(* IEC 61131-3 sources: PortalRobot/Portal_robot/Device/application/FB (part 6) *)

(* ---- FB_TWO_PALLET.st ---- *)
FUNCTION_BLOCK FB_TWO_PALLET
VAR_INPUT
	xSelected : BOOL;
	xManual : BOOL;
	xSafe : BOOL;
	xRobotSwapWindow : BOOL; // Завершено последнее обслуживание: разрешён автоматический обмен
	xRobotOperation : BOOL; // Текущая или уже выданная операция с этим магазином
	xPointsConfigured : BOOL; // Собственная база магазина нужна для ввода в автомат
	xRobotGeometryReady : BOOL; // Собственная база магазина и поддерживаемый интерфейс робота
	xRobotMagazineReady : BOOL; // Ошибки и геометрия магазина; содержимое не блокирует включение
	xConnection : BOOL; // Heartbeat HMI нужен только для ручных команд
	xStopRequest : BOOL; // Общий Stop прерывает движение, но не отключает неподвижный магазин
	xAutoSwap : BOOL;
	xOtherLoaded : BOOL;
	xActivePalletEditAllowed : BOOL;
	xConfigurationChanged : BOOL;
    xIoPneumaticOverride : BOOL; // Прямое воздействие на катушки снимает подтверждение расстановки
	xExternalCommandRejected : BOOL;
	Command : ST_TWO_PALLET_COMMAND;
	Config : ST_TWO_PALLET_CONFIG;
	Input : ST_TWO_PALLET_INPUT;
END_VAR
VAR_OUTPUT
	Status : ST_TWO_PALLET_STATUS;
	Diag : ST_TWO_PALLET_DIAG;
	Error : ST_TWO_PALLET_ERRORS;
	Output : ST_TWO_PALLET_OUTPUT;
END_VAR
VAR
	ePreviousState : E_TWO_PALLET_STATE := E_TWO_PALLET_STATE.IDLE;
	uiFrom : UINT;
	uiTo : UINT;
	uiSelected : UINT;
	uiCandidate : UINT;
	uiPreviousCandidate : UINT;
	uiConfirmedCandidate : UINT;
	uiManualSelected : UINT;
	uiJogDirection : UINT;
	uiSignals : UINT;
	uiSelectedSignals : UINT;
	uiTargetSignals : UINT;
	xPreviousBaseValid : BOOL;
	xConfigValid : BOOL;
	xContradiction : BOOL;
	xPairValid : BOOL;
	xWork : BOOL;
	xExchange : BOOL;
	xIdle : BOOL;
	xBase : BOOL;
	xManualSetupAllowed : BOOL;
	xRecovery : BOOL;
	xPneumaticBase : BOOL;
	xPneumaticRecovery : BOOL;
	xManualPneumaticState : BOOL;
	xAutomaticState : BOOL;
	xAxisMotionState : BOOL;
	xManualState : BOOL;
	xEnableBaseAllowed : BOOL;
	xAutoSwapAllowed : BOOL;
	xExchangeStartedManual : BOOL; // Обмен начат в ручном режиме: без проверки роботной зоны/точек
	xCommandPresent : BOOL;
	xAccepted : BOOL;
	xStateEntry : BOOL;
	xSeenMotion : BOOL;
	xSeenDone : BOOL;
	xLiftUpCommand : BOOL;
	xLiftDownCommand : BOOL;
	xSelectCommand : BOOL;
	xManualLockCommand : BOOL;
	xManualStopCommand : BOOL;
	xManualLockOutTarget : BOOL;
	xManualStopOutTarget : BOOL;
	xLockOutTarget : BOOL;
	xStopOutTarget : BOOL;
	xStartupInitialized : BOOL;
	xTrustedAtScanStart : BOOL;
	lrWork : LREAL;
	lrTarget : LREAL;
	lrSpan : LREAL;
	rTravel : REAL;
	tStateLimit : TIME;
	tonState : TON;
	tonCoil : TON;
	tonJogLease : TON;
	dwPreviousError : DWORD;
END_VAR
VAR CONSTANT
	ERR_DRIVE : DWORD := DWORD#16#100;
	ERR_SENSOR_CONTRADICTION : DWORD := DWORD#16#200;
	ERR_CYLINDER_TIMEOUT : DWORD := DWORD#16#400;
	ERR_MOTION_TIMEOUT : DWORD := DWORD#16#800;
	ERR_LOGIC : DWORD := DWORD#16#1000;
	ERR_SEQUENCE_INTERRUPTED : DWORD := DWORD#16#2000;
	WRN_COMMAND_REJECTED : UINT := UINT#30;
	WRN_ENABLE_POINTS : UINT := UINT#18; // Общий код с FB_MAGAZINE для отсутствующей базы
	WRN_START_REJECTED_BY_OPERATOR : UINT := UINT#31;
	JOG_POSITIVE : UINT := UINT#1;
	JOG_NEGATIVE : UINT := UINT#2;
END_VAR

// --- BEGIN IMPLEMENTATION ---

// Шаги, разрешения и подтверждение положения не восстанавливаются после старта PLC.
IF NOT xStartupInitialized THEN
	Diag.eState := E_TWO_PALLET_STATE.IDLE;
	ePreviousState := E_TWO_PALLET_STATE.IDLE;
	Status.xConfirmed := FALSE;
	Status.xEnabled := FALSE;
	xStartupInitialized := TRUE;
END_IF;

Status.xCompleted := FALSE;
Status.Input := Input;
xTrustedAtScanStart := Status.xConfirmed;

// Все выходные команды импульсные или формируются заново на каждом скане.
Output.xPowerOn := FALSE;
Output.xPowerOff := FALSE;
Output.xDriveReset := FALSE;
Output.xHome := FALSE;
Output.xMove := FALSE;
Output.xStop := FALSE;
Output.xJogPositive := FALSE;
Output.xJogNegative := FALSE;
Output.xTeachOperator := FALSE;
Output.xTeachWork := FALSE;
xLiftUpCommand := FALSE;
xLiftDownCommand := FALSE;
xSelectCommand := FALSE;
xManualLockCommand := FALSE;
xManualStopCommand := FALSE;

// Конфигурация механизма.
xConfigValid := Config.xConfigured
	AND Config.xSignalPatternsConfigured
	AND IsSignalConfigurationValid(uiP1Signals := Config.uiP1Signals, uiP2Signals := Config.uiP2Signals)
	AND (Config.lrTolerance > 0.0)
	AND (Config.lrTolerance <= 20.0)
	AND (ABS(Config.lrWorkP1 - Config.lrExchange) > 2.0 * Config.lrTolerance)
	AND (ABS(Config.lrWorkP2 - Config.lrExchange) > 2.0 * Config.lrTolerance)
	AND ((Config.lrWorkP1 - Config.lrExchange) * (Config.lrWorkP2 - Config.lrExchange) > 0.0)
	AND (Config.lrVelocity > 0.0)
	AND (Config.lrAcceleration > 0.0)
	AND (Config.lrDeceleration > 0.0)
	AND (Config.lrJerk > 0.0)
	AND (Config.tPulse >= T#50MS)
	AND (Config.tCylinder > Config.tPulse)
	AND (Config.tMove > T#0S)
	AND (Config.tHome > T#0S);
Status.xConfigValid := xConfigValid;

// Фактическое состояние пневматики и каретки.
xContradiction := (Input.xLiftUp AND Input.xLiftDown)
	OR (Input.xLockIn AND Input.xLockOut)
	OR (Input.xStopIn AND Input.xStopOut)
	OR (Input.xLimitNegative AND Input.xLimitPositive);
xPairValid := (Input.xLockIn XOR Input.xLockOut)
	AND (Input.xStopIn XOR Input.xStopOut);

uiSignals := UINT#0;
IF Input.xLiftDown THEN uiSignals := uiSignals OR UINT#1; END_IF;
IF Input.xLiftUp THEN uiSignals := uiSignals OR UINT#2; END_IF;
IF Input.xLockIn THEN uiSignals := uiSignals OR UINT#4; END_IF;
IF Input.xLockOut THEN uiSignals := uiSignals OR UINT#8; END_IF;
IF Input.xStopIn THEN uiSignals := uiSignals OR UINT#16; END_IF;
IF Input.xStopOut THEN uiSignals := uiSignals OR UINT#32; END_IF;

uiSelected := UINT#0;
IF xPairValid THEN
	IF (uiSignals AND UINT#60) = (Config.uiP1Signals AND UINT#60) THEN
		uiSelected := UINT#1;
	ELSIF (uiSignals AND UINT#60) = (Config.uiP2Signals AND UINT#60) THEN
		uiSelected := UINT#2;
	END_IF;
END_IF;
xPairValid := xPairValid AND (uiSelected <> UINT#0);

lrWork := Config.lrWorkP1;
uiSelectedSignals := Config.uiP1Signals;
IF uiSelected = UINT#2 THEN
	lrWork := Config.lrWorkP2;
	uiSelectedSignals := Config.uiP2Signals;
END_IF;

xWork := xConfigValid
	AND Input.xHomed
	AND Input.xStandstill
	AND xPairValid
	AND (ABS(Input.lrPosition - lrWork) <= Config.lrTolerance);
xExchange := xConfigValid
	AND Input.xHomed
	AND Input.xStandstill
	AND (ABS(Input.lrPosition - Config.lrExchange) <= Config.lrTolerance);

uiCandidate := UINT#0;
IF xWork
	AND (uiSignals = uiSelectedSignals)
	AND NOT xContradiction
	AND NOT Input.xDriveError
	AND NOT Status.xHomeRequired THEN
	uiCandidate := uiSelected;
END_IF;

xIdle := Diag.eState = E_TWO_PALLET_STATE.IDLE;
xAutomaticState := (Diag.eState = E_TWO_PALLET_STATE.AUTO_LOWER)
	OR (Diag.eState = E_TWO_PALLET_STATE.AUTO_MOVE_TO_EXCHANGE)
	OR (Diag.eState = E_TWO_PALLET_STATE.AUTO_SELECT_PALLET)
	OR (Diag.eState = E_TWO_PALLET_STATE.AUTO_MOVE_TO_WORK)
	OR (Diag.eState = E_TWO_PALLET_STATE.AUTO_RAISE);
xAxisMotionState := (Diag.eState = E_TWO_PALLET_STATE.AUTO_MOVE_TO_EXCHANGE)
	OR (Diag.eState = E_TWO_PALLET_STATE.AUTO_MOVE_TO_WORK)
	OR (Diag.eState = E_TWO_PALLET_STATE.MANUAL_MOVE)
	OR (Diag.eState = E_TWO_PALLET_STATE.MANUAL_HOME)
	OR (Diag.eState = E_TWO_PALLET_STATE.MANUAL_JOG);
xManualState := (Diag.eState = E_TWO_PALLET_STATE.MANUAL_LOWER)
	OR (Diag.eState = E_TWO_PALLET_STATE.MANUAL_RAISE)
	OR (Diag.eState = E_TWO_PALLET_STATE.MANUAL_SELECT_PALLET)
	OR (Diag.eState = E_TWO_PALLET_STATE.MANUAL_MOVE)
	OR (Diag.eState = E_TWO_PALLET_STATE.MANUAL_HOME)
	OR (Diag.eState = E_TWO_PALLET_STATE.MANUAL_JOG)
	OR (Diag.eState = E_TWO_PALLET_STATE.MANUAL_LOCK)
	OR (Diag.eState = E_TWO_PALLET_STATE.MANUAL_STOP);
xManualPneumaticState := (Diag.eState = E_TWO_PALLET_STATE.MANUAL_LOWER)
	OR (Diag.eState = E_TWO_PALLET_STATE.MANUAL_LOCK)
	OR (Diag.eState = E_TWO_PALLET_STATE.MANUAL_STOP);

xBase := xSelected
	AND xConfigValid
	AND Input.xIoMapped
	AND Input.xAxisBound
	AND xSafe
	AND NOT xRobotOperation;
xManualSetupAllowed := xManual
	AND NOT Status.xEnabled
	AND NOT xRobotOperation;
xRecovery := xBase
	AND xManualSetupAllowed
	AND xConnection
	AND xIdle
	AND Input.xStandstill;
xPneumaticBase := xSelected
	AND xManualSetupAllowed
	AND xSafe
	AND Input.xIoMapped
	AND Input.xStandstill;
xPneumaticRecovery := xPneumaticBase AND xIdle;

Status.uiCandidate := uiCandidate;
Status.uiSelected := uiSelected;

// Любое изменение достоверной расстановки аннулирует старое подтверждение.
IF (uiCandidate <> uiPreviousCandidate) OR (xBase <> xPreviousBaseValid) THEN
	Status.udiRevision := Status.udiRevision + UDINT#1;
	IF Status.udiRevision = UDINT#0 THEN
		Status.udiRevision := UDINT#1;
	END_IF;
END_IF;
uiPreviousCandidate := uiCandidate;
xPreviousBaseValid := xBase;

IF xConfigurationChanged THEN
	Status.xConfirmed := FALSE;
	Status.xEnabled := FALSE;
	Status.udiRevision := Status.udiRevision + UDINT#1;
	IF Status.udiRevision = UDINT#0 THEN
		Status.udiRevision := UDINT#1;
	END_IF;
END_IF;

IF xIoPneumaticOverride THEN
    Status.xConfirmed := FALSE;
    Status.xEnabled := FALSE;
    Status.udiRevision := Status.udiRevision + UDINT#1;
    IF Status.udiRevision = UDINT#0 THEN Status.udiRevision := UDINT#1; END_IF;
END_IF;

IF NOT xSelected
	OR NOT xSafe
	OR NOT Input.xAxisBound
	OR NOT Input.xIoMapped
	OR NOT xConfigValid
	OR Input.xDriveError
	OR NOT Input.xPowered
	OR (xIdle AND (uiCandidate <> uiConfirmedCandidate)) THEN
	Status.xConfirmed := FALSE;
END_IF;
// Первая невыполненная предпосылка для HMI.
Diag.uiReason := UINT#0;
IF NOT xSelected THEN
	Diag.uiReason := UINT#1;
ELSIF NOT xConfigValid THEN
	Diag.uiReason := UINT#2;
ELSIF NOT Input.xAxisBound OR NOT Input.xIoMapped THEN
	Diag.uiReason := UINT#3;
ELSIF NOT xSafe THEN
	Diag.uiReason := UINT#4;
ELSIF NOT xConnection THEN
	Diag.uiReason := UINT#17;
ELSIF Input.xDriveError THEN
	Diag.uiReason := UINT#6;
ELSIF Error.dwErrorActive <> DWORD#0 THEN
	Diag.uiReason := UINT#19;
ELSIF NOT Input.xPowered THEN
	Diag.uiReason := UINT#18;
ELSIF xContradiction THEN
	Diag.uiReason := UINT#7;
ELSIF Status.xHomeRequired OR NOT Input.xHomed THEN
	Diag.uiReason := UINT#8;
ELSIF NOT xPairValid THEN
	Diag.uiReason := UINT#9;
ELSIF NOT Input.xStandstill THEN
	Diag.uiReason := UINT#10;
ELSIF NOT xWork THEN
	Diag.uiReason := UINT#11;
ELSIF uiSignals <> uiSelectedSignals THEN
	Diag.uiReason := UINT#12;
ELSIF NOT xIdle THEN
	Diag.uiReason := UINT#22;
ELSIF xRobotOperation THEN
	Diag.uiReason := UINT#5;
ELSIF xManual AND Status.xEnabled THEN
	Diag.uiReason := UINT#21;
ELSIF NOT xManual AND NOT xRobotSwapWindow THEN
	Diag.uiReason := UINT#23;
ELSIF NOT xRobotMagazineReady THEN
	Diag.uiReason := UINT#16;
ELSIF NOT xPointsConfigured THEN
	Diag.uiReason := UINT#15;
ELSIF NOT Status.xConfirmed AND NOT xManual THEN
	Diag.uiReason := UINT#20;
ELSIF NOT Status.xConfirmed THEN
	Diag.uiReason := UINT#13;
END_IF;

// Аварии механизма: биты 8..13 зарезервированы в MAGAZINE_LOGIC_1/2.
IF xSelected AND Input.xDriveError THEN
	Error.dwErrorActive := Error.dwErrorActive OR ERR_DRIVE;
	Status.xHomeRequired := TRUE;
END_IF;

IF xSelected AND xContradiction THEN
	Error.dwErrorActive := Error.dwErrorActive OR ERR_SENSOR_CONTRADICTION;
END_IF;

IF xSelected
	AND NOT xIdle
	AND (((NOT xBase) AND NOT (xManualPneumaticState AND xPneumaticBase))
		OR (xManualState AND NOT xManual)
		OR ((NOT xConnection) AND xManualState AND NOT xManualPneumaticState) OR xStopRequest
		OR (xAutomaticState AND ((xExchangeStartedManual AND NOT xManual)
			OR (NOT xExchangeStartedManual AND NOT xRobotSwapWindow)))) THEN
	Error.dwErrorActive := Error.dwErrorActive OR ERR_SEQUENCE_INTERRUPTED;
	Diag.eState := E_TWO_PALLET_STATE.IDLE;
	Output.xStop := TRUE;
END_IF;

IF xSelected AND (xTrustedAtScanStart OR xAutomaticState) THEN
	IF ((Diag.eState <> E_TWO_PALLET_STATE.AUTO_SELECT_PALLET) AND NOT xPairValid)
		OR (((Diag.eState = E_TWO_PALLET_STATE.AUTO_MOVE_TO_EXCHANGE)
			OR (Diag.eState = E_TWO_PALLET_STATE.AUTO_MOVE_TO_WORK))
			AND (NOT Input.xLiftDown OR Input.xLiftUp))
		OR (xIdle AND (uiCandidate = UINT#0)) THEN
		Error.dwErrorActive := Error.dwErrorActive OR ERR_LOGIC;
	END_IF;
END_IF;

IF xSelected
	AND xTrustedAtScanStart
	AND (NOT xSafe
		OR NOT Input.xAxisBound
		OR NOT Input.xIoMapped
		OR NOT Input.xPowered) THEN
	Error.dwErrorActive := Error.dwErrorActive OR ERR_SEQUENCE_INTERRUPTED;
END_IF;

IF xSelected
	AND ((xContradiction AND NOT xIdle AND NOT xManualPneumaticState)
		OR (Input.xDriveError AND xAxisMotionState)) THEN
	Diag.eState := E_TWO_PALLET_STATE.IDLE;
	Output.xStop := TRUE;
END_IF;

IF xSelected AND NOT Input.xPowered AND (xAutomaticState OR xAxisMotionState) THEN
	Error.dwErrorActive := Error.dwErrorActive OR ERR_SEQUENCE_INTERRUPTED;
	Status.xHomeRequired := TRUE;
	Diag.eState := E_TWO_PALLET_STATE.IDLE;
	Output.xStop := TRUE;
END_IF;

IF Error.dwErrorActive <> DWORD#0 THEN
	Status.xEnabled := FALSE;
	Status.xConfirmed := FALSE;
	IF xAutomaticState THEN
		Diag.eState := E_TWO_PALLET_STATE.IDLE;
		Output.xStop := TRUE;
	END_IF;
END_IF;

// Разрешения считаются только владельцем механизма.
Status.xConfirmAllowed := xRecovery
	AND Input.xPowered
	AND (uiCandidate <> UINT#0)
	AND (Error.dwErrorActive = DWORD#0);
Status.xStartAllowed := Status.xConfirmAllowed
	AND xRobotMagazineReady
	AND xPointsConfigured;
// Включение подтверждённого магазина не двигает палету и не снимает резерв
// возврата изделия. Иначе Disable при грузе в роботе блокирует продолжение цикла.
// Общая технологическая готовность не зависит от heartbeat HMI.
xEnableBaseAllowed := xBase
	AND xIdle
	AND Status.xConfirmed
	AND xRobotMagazineReady
	AND xPointsConfigured
	AND (uiCandidate = Status.uiRobotPallet)
	AND Input.xPowered
	AND (Error.dwErrorActive = DWORD#0);
Status.xEnableAllowed := xEnableBaseAllowed AND xConnection;
// Обмен не требует глобальной остановки робота: проверяется только отсутствие
// текущей или уже выданной операции именно с этим магазином.
Status.xSwapAllowed := xBase
	AND xConnection
	AND xIdle
	AND Input.xStandstill
	AND Input.xPowered
	AND (Error.dwErrorActive = DWORD#0)
	AND Status.xConfirmed
	AND (uiCandidate = Status.uiRobotPallet)
	AND NOT Status.xEnabled
	AND NOT xStopRequest
	AND (xRobotSwapWindow OR xManual);
xAutoSwapAllowed := xEnableBaseAllowed
	AND xRobotSwapWindow
	AND Status.xEnabled
	AND xOtherLoaded;
Status.xPowerAllowed := xRecovery
	AND NOT Input.xDriveError
	AND NOT xContradiction;
Status.xDriveResetAllowed := xSelected
	AND xManualSetupAllowed
	AND xConnection
	AND Input.xAxisBound
	AND Input.xStandstill
	AND xIdle;
Status.xLowerAllowed := xPneumaticRecovery;
Status.xRaiseAllowed := xRecovery
	AND NOT xContradiction
	AND NOT Status.xHomeRequired;
Status.xSelectAllowed := xRecovery
	AND NOT xContradiction
	AND Input.xLiftDown
	AND NOT Input.xLiftUp
	AND xExchange;
// Наладочные команды замка и фиксатора независимы от подъёма и координаты.
// Это позволяет вернуть герконы в согласованное состояние после остановки.
Status.xLockAllowed := xPneumaticRecovery;
Status.xStopAllowed := xPneumaticRecovery;
Status.xHomeAllowed := xRecovery
	AND Input.xPowered
	AND NOT Input.xDriveError
	AND Input.xLiftDown
	AND NOT Input.xLiftUp
	AND xPairValid
	AND NOT xContradiction;
Status.xMoveAllowed := Status.xHomeAllowed
	AND Input.xHomed
	AND NOT Status.xHomeRequired;
Status.xJogAllowed := Status.xHomeAllowed;
Status.xTeachOperatorAllowed := Status.xMoveAllowed
	AND Input.xLiftDown
	AND NOT Input.xLiftUp;
Status.xTeachWorkAllowed := Status.xTeachOperatorAllowed
	AND ((uiSelected = UINT#1) OR (uiSelected = UINT#2));
Status.xResetAllowed := xRecovery
	AND (Error.dwErrorActive <> DWORD#0)
	AND NOT xContradiction
	AND NOT Input.xDriveError
	AND NOT Status.xHomeRequired
	AND xPairValid
	AND (Input.xLiftDown XOR Input.xLiftUp);
Status.xConfigAllowed := xSelected
	AND xManualSetupAllowed
	AND xIdle
	AND NOT Status.xEnabled
	AND (Input.xStandstill OR NOT Input.xAxisBound)
	AND NOT Input.xPowered;

// Командный интерфейс FB не зависит от транспортных номеров HMI 1..19.
xCommandPresent := Command.xEnable
	OR Command.xConfirm
	OR Command.xStart
	OR Command.xRejectStart
	OR Command.xDisable
	OR Command.xSwap
	OR Command.xPowerOn
	OR Command.xPowerOff
	OR Command.xDriveReset
	OR Command.xHome
	OR Command.xLower
	OR Command.xRaise
	OR Command.xSelectPallet
	OR Command.xLockIn
	OR Command.xLockOut
	OR Command.xStopIn
	OR Command.xStopOut
	OR Command.xMoveToExchange
	OR Command.xMoveToWork
	OR Command.xStop
	OR Command.xReset
	OR Command.xJogPositive
	OR Command.xJogNegative
	OR Command.xJogRelease
	OR Command.xTeachOperator
	OR Command.xTeachWork;
xAccepted := NOT xCommandPresent;

IF Command.xStart THEN
	IF Status.xStartAllowed
		AND (Command.udiRevision = Status.udiRevision)
		AND (Command.uiPallet = uiCandidate) THEN
		Status.uiRobotPallet := uiCandidate;
		uiConfirmedCandidate := uiCandidate;
		Status.xConfirmed := TRUE;
		Status.xEnabled := TRUE;
		Status.rP1 := 0.0;
		Status.rP2 := 0.0;
		IF uiCandidate = UINT#1 THEN
			Status.rP1 := 1.0;
		ELSE
			Status.rP2 := 1.0;
		END_IF;
		xAccepted := TRUE;
	END_IF;
ELSIF Command.xRejectStart THEN
	Diag.stWarning.uiCode := WRN_START_REJECTED_BY_OPERATOR;
	Diag.stWarning.udiSequence := Diag.stWarning.udiSequence + UDINT#1;
	IF Diag.stWarning.udiSequence = UDINT#0 THEN
		Diag.stWarning.udiSequence := UDINT#1;
	END_IF;
	xAccepted := TRUE;
ELSIF Command.xEnable THEN
	IF Status.xEnableAllowed THEN
		Status.xEnabled := TRUE;
		xAccepted := TRUE;
	END_IF;
ELSIF Command.xConfirm THEN
	IF Status.xConfirmAllowed
		AND (Command.udiRevision = Status.udiRevision)
		AND (Command.uiPallet = uiCandidate) THEN
		Status.uiRobotPallet := uiCandidate;
		uiConfirmedCandidate := uiCandidate;
		Status.xConfirmed := TRUE;
		Status.rP1 := 0.0;
		Status.rP2 := 0.0;
		IF uiCandidate = UINT#1 THEN
			Status.rP1 := 1.0;
		ELSE
			Status.rP2 := 1.0;
		END_IF;
		xAccepted := TRUE;
	END_IF;
ELSIF Command.xDisable THEN
	Status.xEnabled := FALSE;
	xAccepted := TRUE;
ELSIF Command.xSwap THEN
	IF Status.xSwapAllowed THEN
		xExchangeStartedManual := xManual;
		Diag.eState := E_TWO_PALLET_STATE.AUTO_LOWER;
		xAccepted := TRUE;
	END_IF;
ELSIF Command.xPowerOn THEN
	IF Status.xPowerAllowed THEN
		Output.xPowerOn := TRUE;
		xAccepted := TRUE;
	END_IF;
ELSIF Command.xPowerOff THEN
	IF Status.xDriveResetAllowed THEN
		Output.xPowerOff := TRUE;
		Status.xConfirmed := FALSE;
		Status.xEnabled := FALSE;
		xAccepted := TRUE;
	END_IF;
ELSIF Command.xDriveReset THEN
	IF Status.xDriveResetAllowed AND Input.xDriveError THEN
		Output.xDriveReset := TRUE;
		Status.xConfirmed := FALSE;
		Status.xEnabled := FALSE;
		Status.xHomeRequired := TRUE;
		xAccepted := TRUE;
	END_IF;
ELSIF Command.xHome THEN
	IF Status.xHomeAllowed THEN
		Diag.eState := E_TWO_PALLET_STATE.MANUAL_HOME;
		xAccepted := TRUE;
	END_IF;
ELSIF Command.xLower THEN
	IF Status.xLowerAllowed THEN
		Diag.eState := E_TWO_PALLET_STATE.MANUAL_LOWER;
		xAccepted := TRUE;
	END_IF;
ELSIF Command.xRaise THEN
	IF Status.xRaiseAllowed THEN
		Diag.eState := E_TWO_PALLET_STATE.MANUAL_RAISE;
		xAccepted := TRUE;
	END_IF;
ELSIF Command.xSelectPallet THEN
	IF Status.xSelectAllowed
		AND ((Command.uiPallet = UINT#1) OR (Command.uiPallet = UINT#2)) THEN
		uiTo := Command.uiPallet;
		Diag.eState := E_TWO_PALLET_STATE.MANUAL_SELECT_PALLET;
		xAccepted := TRUE;
	END_IF;
ELSIF Command.xLockIn OR Command.xLockOut THEN
	IF Status.xLockAllowed THEN
		xManualLockOutTarget := Command.xLockOut;
		Diag.eState := E_TWO_PALLET_STATE.MANUAL_LOCK;
		xAccepted := TRUE;
	END_IF;
ELSIF Command.xStopIn OR Command.xStopOut THEN
	IF Status.xStopAllowed THEN
		xManualStopOutTarget := Command.xStopOut;
		Diag.eState := E_TWO_PALLET_STATE.MANUAL_STOP;
		xAccepted := TRUE;
	END_IF;
ELSIF Command.xMoveToExchange OR Command.xMoveToWork THEN
	IF Status.xMoveAllowed THEN
		lrTarget := Config.lrExchange;
		IF Command.xMoveToWork THEN
			lrTarget := lrWork;
		END_IF;
		Diag.eState := E_TWO_PALLET_STATE.MANUAL_MOVE;
		xAccepted := TRUE;
	END_IF;
ELSIF Command.xStop THEN
	Status.xEnabled := FALSE;
	// Stop неподвижного механизма не является ручным вмешательством.
	IF (Diag.eState <> E_TWO_PALLET_STATE.IDLE) OR (Input.xPowered AND NOT Input.xStandstill) THEN
		Output.xStop := TRUE;
		Status.xConfirmed := FALSE;
		Error.dwErrorActive := Error.dwErrorActive OR ERR_SEQUENCE_INTERRUPTED;
	END_IF;
	Diag.eState := E_TWO_PALLET_STATE.IDLE;
	uiJogDirection := UINT#0;
	xAccepted := TRUE;
ELSIF Command.xReset THEN
	IF Status.xResetAllowed THEN
		Error.dwErrorLast := Error.dwErrorActive;
		Error.dwErrorActive := DWORD#0;
		Status.xConfirmed := FALSE;
		Status.xEnabled := FALSE;
		xAccepted := TRUE;
	END_IF;
ELSIF Command.xJogPositive OR Command.xJogNegative THEN
	IF Status.xJogAllowed
		OR ((Diag.eState = E_TWO_PALLET_STATE.MANUAL_JOG)
			AND xBase
			AND xManualSetupAllowed
			AND xConnection) THEN
		Diag.eState := E_TWO_PALLET_STATE.MANUAL_JOG;
		IF Command.xJogPositive THEN
			uiJogDirection := JOG_POSITIVE;
		ELSE
			uiJogDirection := JOG_NEGATIVE;
		END_IF;
		xAccepted := TRUE;
	END_IF;
ELSIF Command.xJogRelease THEN
	uiJogDirection := UINT#0;
	IF Diag.eState = E_TWO_PALLET_STATE.MANUAL_JOG THEN
		Diag.eState := E_TWO_PALLET_STATE.IDLE;
		Output.xStop := TRUE;
	END_IF;
	xAccepted := TRUE;
ELSIF Command.xTeachOperator THEN
	IF Status.xTeachOperatorAllowed THEN
		Output.xTeachOperator := TRUE;
		xAccepted := TRUE;
	END_IF;
ELSIF Command.xTeachWork THEN
	IF Status.xTeachWorkAllowed THEN
		Output.xTeachWork := TRUE;
		xAccepted := TRUE;
	END_IF;
END_IF;

IF xCommandPresent AND NOT xAccepted THEN
	IF (Command.xEnable OR Command.xStart) AND NOT xPointsConfigured THEN
		Diag.stWarning.uiCode := WRN_ENABLE_POINTS;
	ELSE
		Diag.stWarning.uiCode := WRN_COMMAND_REJECTED;
	END_IF;
	Diag.stWarning.udiSequence := Diag.stWarning.udiSequence + UDINT#1;
	IF Diag.stWarning.udiSequence = UDINT#0 THEN
		Diag.stWarning.udiSequence := UDINT#1;
	END_IF;
END_IF;

IF xExternalCommandRejected THEN
	Diag.stWarning.uiCode := WRN_COMMAND_REJECTED;
	Diag.stWarning.udiSequence := Diag.stWarning.udiSequence + UDINT#1;
	IF Diag.stWarning.udiSequence = UDINT#0 THEN
		Diag.stWarning.udiSequence := UDINT#1;
	END_IF;
END_IF;

Status.xCommandAccepted := xAccepted;

IF xAutoSwap
	AND xAutoSwapAllowed
	AND NOT Output.xStop
	AND NOT xCommandPresent THEN
	xExchangeStartedManual := FALSE;
	Diag.eState := E_TWO_PALLET_STATE.AUTO_LOWER;
END_IF;

// Стоп ячейки имеет приоритет над командой, принятой в том же скане.
// В IDLE при остановленной оси сохраняем включение и подтверждение.
// Собственные Command.xStop / Command.xDisable отдельно отключают магазин.
IF xStopRequest THEN
	IF (Diag.eState <> E_TWO_PALLET_STATE.IDLE) OR (Input.xPowered AND NOT Input.xStandstill) THEN
		Error.dwErrorActive := Error.dwErrorActive OR ERR_SEQUENCE_INTERRUPTED;
		Output.xStop := TRUE;
		Status.xConfirmed := FALSE;
		Status.xEnabled := FALSE;
	END_IF;
	Diag.eState := E_TWO_PALLET_STATE.IDLE;
END_IF;

// Команда могла сменить состояние в этом же скане — обновляем классификацию
// до обработки входа в шаг и запуска таймеров.
xAutomaticState := (Diag.eState = E_TWO_PALLET_STATE.AUTO_LOWER)
	OR (Diag.eState = E_TWO_PALLET_STATE.AUTO_MOVE_TO_EXCHANGE)
	OR (Diag.eState = E_TWO_PALLET_STATE.AUTO_SELECT_PALLET)
	OR (Diag.eState = E_TWO_PALLET_STATE.AUTO_MOVE_TO_WORK)
	OR (Diag.eState = E_TWO_PALLET_STATE.AUTO_RAISE);
xManualState := (Diag.eState = E_TWO_PALLET_STATE.MANUAL_LOWER)
	OR (Diag.eState = E_TWO_PALLET_STATE.MANUAL_RAISE)
	OR (Diag.eState = E_TWO_PALLET_STATE.MANUAL_SELECT_PALLET)
	OR (Diag.eState = E_TWO_PALLET_STATE.MANUAL_MOVE)
	OR (Diag.eState = E_TWO_PALLET_STATE.MANUAL_HOME)
	OR (Diag.eState = E_TWO_PALLET_STATE.MANUAL_JOG)
	OR (Diag.eState = E_TWO_PALLET_STATE.MANUAL_LOCK)
	OR (Diag.eState = E_TWO_PALLET_STATE.MANUAL_STOP);
xManualPneumaticState := (Diag.eState = E_TWO_PALLET_STATE.MANUAL_LOWER)
	OR (Diag.eState = E_TWO_PALLET_STATE.MANUAL_LOCK)
	OR (Diag.eState = E_TWO_PALLET_STATE.MANUAL_STOP);

IF (Diag.eState = E_TWO_PALLET_STATE.AUTO_LOWER)
	AND (ePreviousState <> E_TWO_PALLET_STATE.AUTO_LOWER) THEN
	uiFrom := Status.uiRobotPallet;
	uiTo := UINT#3 - uiFrom;
END_IF;

xStateEntry := Diag.eState <> ePreviousState;
IF xManualState AND xStateEntry THEN
	Status.xConfirmed := FALSE;
	Status.xEnabled := FALSE;
	Status.udiRevision := Status.udiRevision + UDINT#1;
	IF Status.udiRevision = UDINT#0 THEN
		Status.udiRevision := UDINT#1;
	END_IF;
END_IF;

IF xStateEntry THEN
	xSeenMotion := FALSE;
	xSeenDone := FALSE;
	IF (Diag.eState = E_TWO_PALLET_STATE.MANUAL_MOVE)
		OR (Diag.eState = E_TWO_PALLET_STATE.MANUAL_HOME)
		OR (Diag.eState = E_TWO_PALLET_STATE.MANUAL_JOG) THEN
		uiManualSelected := uiSelected;
	END_IF;
ELSIF Input.xMotionDone THEN
	xSeenDone := TRUE;
END_IF;

IF NOT Input.xStandstill THEN
	xSeenMotion := TRUE;
END_IF;

tStateLimit := Config.tCylinder;
IF (Diag.eState = E_TWO_PALLET_STATE.AUTO_MOVE_TO_EXCHANGE)
	OR (Diag.eState = E_TWO_PALLET_STATE.AUTO_MOVE_TO_WORK)
	OR (Diag.eState = E_TWO_PALLET_STATE.MANUAL_MOVE) THEN
	tStateLimit := Config.tMove;
END_IF;
IF Diag.eState = E_TWO_PALLET_STATE.MANUAL_HOME THEN
	tStateLimit := Config.tHome;
END_IF;

tonState(
	IN := NOT xIdle
		AND (Diag.eState <> E_TWO_PALLET_STATE.MANUAL_JOG)
		AND NOT xStateEntry,
	PT := tStateLimit);
tonCoil(
	IN := NOT xIdle AND NOT xStateEntry,
	PT := Config.tPulse);
tonJogLease(
	IN := (Diag.eState = E_TWO_PALLET_STATE.MANUAL_JOG)
		AND NOT (Command.xJogPositive OR Command.xJogNegative),
	PT := T#350MS);
ePreviousState := Diag.eState;

// Автомат обмена и ручного восстановления.
uiTargetSignals := Config.uiP1Signals;
IF uiTo = UINT#2 THEN uiTargetSignals := Config.uiP2Signals; END_IF;
CASE Diag.eState OF
	E_TWO_PALLET_STATE.AUTO_LOWER,
	E_TWO_PALLET_STATE.MANUAL_LOWER:
		xLiftDownCommand := TRUE;
		IF Input.xLiftDown AND NOT Input.xLiftUp THEN
			IF Diag.eState = E_TWO_PALLET_STATE.AUTO_LOWER THEN
				Diag.eState := E_TWO_PALLET_STATE.AUTO_MOVE_TO_EXCHANGE;
				lrTarget := Config.lrExchange;
			ELSE
				Diag.eState := E_TWO_PALLET_STATE.IDLE;
			END_IF;
		END_IF;

	E_TWO_PALLET_STATE.AUTO_MOVE_TO_EXCHANGE,
	E_TWO_PALLET_STATE.AUTO_MOVE_TO_WORK,
	E_TWO_PALLET_STATE.MANUAL_MOVE:
		IF Diag.eState = E_TWO_PALLET_STATE.AUTO_MOVE_TO_WORK THEN
			lrTarget := Config.lrWorkP1;
			IF uiTo = UINT#2 THEN
				lrTarget := Config.lrWorkP2;
			END_IF;
		END_IF;

		IF NOT Input.xLiftDown
			OR Input.xLiftUp
			OR NOT xPairValid
			OR Status.xHomeRequired
			OR ((Diag.eState = E_TWO_PALLET_STATE.AUTO_MOVE_TO_EXCHANGE) AND (uiSelected <> uiFrom))
			OR ((Diag.eState = E_TWO_PALLET_STATE.AUTO_MOVE_TO_WORK) AND (uiSelected <> uiTo))
			OR ((Diag.eState = E_TWO_PALLET_STATE.MANUAL_MOVE) AND (uiSelected <> uiManualSelected))
			OR (Input.xLimitPositive AND (lrTarget > Input.lrPosition + Config.lrTolerance))
			OR (Input.xLimitNegative AND (lrTarget < Input.lrPosition - Config.lrTolerance)) THEN
			Error.dwErrorActive := Error.dwErrorActive OR ERR_LOGIC;
			Diag.eState := E_TWO_PALLET_STATE.IDLE;
			Output.xStop := TRUE;
		ELSE
			Output.lrTarget := lrTarget;
			Output.xMove := xStateEntry;
			IF Input.xStandstill
				AND (ABS(Input.lrPosition - lrTarget) <= Config.lrTolerance)
				AND ((xSeenMotion OR xSeenDone) OR xStateEntry) THEN
				Output.xMove := FALSE;
				IF Diag.eState = E_TWO_PALLET_STATE.AUTO_MOVE_TO_EXCHANGE THEN
					Diag.eState := E_TWO_PALLET_STATE.AUTO_SELECT_PALLET;
				ELSIF Diag.eState = E_TWO_PALLET_STATE.AUTO_MOVE_TO_WORK THEN
					Diag.eState := E_TWO_PALLET_STATE.AUTO_RAISE;
				ELSE
					Diag.eState := E_TWO_PALLET_STATE.IDLE;
				END_IF;
			END_IF;
		END_IF;

	E_TWO_PALLET_STATE.AUTO_SELECT_PALLET,
	E_TWO_PALLET_STATE.MANUAL_SELECT_PALLET:
		IF NOT xExchange OR NOT Input.xLiftDown OR Input.xLiftUp THEN
			Error.dwErrorActive := Error.dwErrorActive OR ERR_LOGIC;
			Diag.eState := E_TWO_PALLET_STATE.IDLE;
			Output.xStop := TRUE;
		ELSE
			xSelectCommand := TRUE;
		END_IF;
		IF (uiSelected = uiTo) AND xPairValid AND NOT Output.xStop THEN
			IF Diag.eState = E_TWO_PALLET_STATE.AUTO_SELECT_PALLET THEN
				Diag.eState := E_TWO_PALLET_STATE.AUTO_MOVE_TO_WORK;
			ELSE
				Diag.eState := E_TWO_PALLET_STATE.IDLE;
			END_IF;
		END_IF;

	E_TWO_PALLET_STATE.MANUAL_LOCK:
		IF xManualLockOutTarget THEN
			xManualLockCommand := NOT Input.xLockOut OR Input.xLockIn;
			IF Input.xLockOut AND NOT Input.xLockIn THEN Diag.eState := E_TWO_PALLET_STATE.IDLE; END_IF;
		ELSE
			xManualLockCommand := NOT Input.xLockIn OR Input.xLockOut;
			IF Input.xLockIn AND NOT Input.xLockOut THEN Diag.eState := E_TWO_PALLET_STATE.IDLE; END_IF;
		END_IF;

	E_TWO_PALLET_STATE.MANUAL_STOP:
		IF xManualStopOutTarget THEN
			xManualStopCommand := NOT Input.xStopOut OR Input.xStopIn;
			IF Input.xStopOut AND NOT Input.xStopIn THEN Diag.eState := E_TWO_PALLET_STATE.IDLE; END_IF;
		ELSE
			xManualStopCommand := NOT Input.xStopIn OR Input.xStopOut;
			IF Input.xStopIn AND NOT Input.xStopOut THEN Diag.eState := E_TWO_PALLET_STATE.IDLE; END_IF;
		END_IF;

	E_TWO_PALLET_STATE.AUTO_RAISE:
		// Завершение обмена устанавливает подъём по выбранной конфигурации
		// только после фактического останова в рабочей позиции.
		IF NOT xWork
			OR Status.xHomeRequired
			OR (uiSelected <> uiTo) THEN
			Error.dwErrorActive := Error.dwErrorActive OR ERR_LOGIC;
			Diag.eState := E_TWO_PALLET_STATE.IDLE;
			Output.xStop := TRUE;
		ELSE
			xLiftUpCommand := (uiTargetSignals AND UINT#2) <> UINT#0;
			xLiftDownCommand := NOT xLiftUpCommand;
			IF uiSignals = uiTargetSignals THEN
				Status.uiRobotPallet := uiTo;
				uiConfirmedCandidate := uiTo;
				Status.xConfirmed := TRUE;
				Status.xCompleted := TRUE;
				Diag.eState := E_TWO_PALLET_STATE.IDLE;
			END_IF;
		END_IF;

	E_TWO_PALLET_STATE.MANUAL_RAISE:
		// Наладочный подъём не требует HOME-координаты или рабочей позиции.
		IF NOT Input.xStandstill OR NOT xManual OR xContradiction OR Status.xHomeRequired THEN
			Error.dwErrorActive := Error.dwErrorActive OR ERR_LOGIC;
			Diag.eState := E_TWO_PALLET_STATE.IDLE;
			Output.xStop := TRUE;
		ELSE
			xLiftUpCommand := TRUE;
			IF Input.xLiftUp AND NOT Input.xLiftDown THEN
				Diag.eState := E_TWO_PALLET_STATE.IDLE;
			END_IF;
		END_IF;

	E_TWO_PALLET_STATE.MANUAL_HOME:
		Output.xHome := xStateEntry;
		IF xSeenDone
			AND Input.xHomed
			AND Input.xStandstill
			AND NOT xStateEntry THEN
			Status.xHomeRequired := FALSE;
			Diag.eState := E_TWO_PALLET_STATE.IDLE;
		END_IF;

	E_TWO_PALLET_STATE.MANUAL_JOG:
		IF tonJogLease.Q OR NOT xConnection OR (uiJogDirection = UINT#0) THEN
			Diag.eState := E_TWO_PALLET_STATE.IDLE;
			Output.xStop := TRUE;
		ELSE
			Output.xJogPositive := (uiJogDirection = JOG_POSITIVE) AND NOT Input.xLimitPositive;
			Output.xJogNegative := (uiJogDirection = JOG_NEGATIVE) AND NOT Input.xLimitNegative;
		END_IF;

	E_TWO_PALLET_STATE.IDLE:
		uiJogDirection := UINT#0;

ELSE
	Error.dwErrorActive := Error.dwErrorActive OR ERR_LOGIC;
	Diag.eState := E_TWO_PALLET_STATE.IDLE;
	Output.xStop := TRUE;
END_CASE;
IF Diag.eState = E_TWO_PALLET_STATE.IDLE THEN xExchangeStartedManual := FALSE; END_IF;

// Низ П2 и выбранное зацепление контролируются всё время Home/JOG.
IF ((Diag.eState = E_TWO_PALLET_STATE.MANUAL_HOME)
	OR (Diag.eState = E_TWO_PALLET_STATE.MANUAL_JOG))
	AND (NOT Input.xLiftDown
		OR Input.xLiftUp
		OR NOT xPairValid
		OR (uiSelected <> uiManualSelected)
		OR xContradiction
		OR Input.xDriveError
		OR NOT Input.xPowered) THEN
	Error.dwErrorActive := Error.dwErrorActive OR ERR_LOGIC;
	Diag.eState := E_TWO_PALLET_STATE.IDLE;
	Output.xStop := TRUE;
END_IF;

IF tonState.Q THEN
	IF (ePreviousState = E_TWO_PALLET_STATE.AUTO_MOVE_TO_EXCHANGE)
		OR (ePreviousState = E_TWO_PALLET_STATE.AUTO_MOVE_TO_WORK)
		OR (ePreviousState = E_TWO_PALLET_STATE.MANUAL_MOVE)
		OR (ePreviousState = E_TWO_PALLET_STATE.MANUAL_HOME) THEN
		Error.dwErrorActive := Error.dwErrorActive OR ERR_MOTION_TIMEOUT;
		Status.xHomeRequired := TRUE;
	ELSE
		Error.dwErrorActive := Error.dwErrorActive OR ERR_CYLINDER_TIMEOUT;
	END_IF;
	Diag.eState := E_TWO_PALLET_STATE.IDLE;
	Output.xStop := TRUE;
END_IF;

IF (((NOT xBase) AND NOT (xManualPneumaticState AND xPneumaticBase))
	OR ((NOT xConnection) AND xManualState AND NOT xManualPneumaticState))
	AND (ePreviousState <> E_TWO_PALLET_STATE.IDLE)
	OR Output.xStop THEN
	Output.xMove := FALSE;
	Output.xHome := FALSE;
	Output.xJogPositive := FALSE;
	Output.xJogNegative := FALSE;
	xLiftUpCommand := FALSE;
	xLiftDownCommand := FALSE;
	xSelectCommand := FALSE;
	xManualLockCommand := FALSE;
	xManualStopCommand := FALSE;
END_IF;

// Автоматический обмен переключает пару совместно; ручное восстановление — каждый цилиндр отдельно.
xLockOutTarget := (uiTargetSignals AND UINT#8) <> UINT#0;
xStopOutTarget := (uiTargetSignals AND UINT#32) <> UINT#0;
Output.xLiftUp := xBase AND xLiftUpCommand AND NOT tonCoil.Q;
Output.xLiftDown := (xBase OR xPneumaticBase) AND xLiftDownCommand AND NOT tonCoil.Q;
Output.xLockOut := (xBase AND xSelectCommand AND xLockOutTarget
	OR xPneumaticBase AND xManualLockCommand AND xManualLockOutTarget) AND NOT tonCoil.Q;
Output.xLockIn := (xBase AND xSelectCommand AND NOT xLockOutTarget
	OR xPneumaticBase AND xManualLockCommand AND NOT xManualLockOutTarget) AND NOT tonCoil.Q;
Output.xStopOut := (xBase AND xSelectCommand AND xStopOutTarget
	OR xPneumaticBase AND xManualStopCommand AND xManualStopOutTarget) AND NOT tonCoil.Q;
Output.xStopIn := (xBase AND xSelectCommand AND NOT xStopOutTarget
	OR xPneumaticBase AND xManualStopCommand AND NOT xManualStopOutTarget) AND NOT tonCoil.Q;

// Поза для 3D — оценка по координате каретки и подтверждённому зацеплению.
IF xPairValid AND Input.xHomed THEN
	lrSpan := lrWork - Config.lrExchange;
	IF ABS(lrSpan) > Config.lrTolerance THEN
		rTravel := LREAL_TO_REAL(
			LIMIT(0.0, (Input.lrPosition - Config.lrExchange) / lrSpan, 1.0));
		IF uiSelected = UINT#1 THEN
			Status.rP1 := rTravel;
		ELSE
			Status.rP2 := rTravel;
		END_IF;
	END_IF;
END_IF;

IF Input.xLiftUp AND NOT Input.xLiftDown THEN
	Status.rLift := 1.0;
ELSIF Input.xLiftDown AND NOT Input.xLiftUp THEN
	Status.rLift := 0.0;
END_IF;

// Диагностика и совместимый публичный Status формируются в одном месте.
IF (Error.dwErrorActive <> dwPreviousError)
	AND (Error.dwErrorActive <> DWORD#0) THEN
	Diag.eFaultState := ePreviousState;
END_IF;
dwPreviousError := Error.dwErrorActive;

IF Error.dwErrorActive <> DWORD#0 THEN
	Error.dwErrorLast := Error.dwErrorActive;
	Status.xConfirmed := FALSE;
	Status.xEnabled := FALSE;
END_IF;
Error.dwAlarmActive := Error.dwErrorActive;
Error.stErrorActive := UpdateErrorView(dwError := Error.dwErrorActive);
Error.stErrorLast := UpdateErrorView(dwError := Error.dwErrorLast);

Status.uiStep := TO_UINT(Diag.eState);
Status.uiFaultStep := TO_UINT(Diag.eFaultState);
Status.uiReason := Diag.uiReason;
Status.dwError := Error.dwErrorActive;
Status.stWarning := Diag.stWarning;
Status.xBusy := Diag.eState <> E_TWO_PALLET_STATE.IDLE;
Status.xError := Error.dwErrorActive <> DWORD#0;

// Команда или автомат могли занять механизм после первоначального расчёта
// разрешений. Не публикуем устаревшее разрешение ещё на один скан.
IF Status.xBusy THEN
	Status.xConfirmAllowed := FALSE;
	Status.xStartAllowed := FALSE;
	Status.xEnableAllowed := FALSE;
	Status.xSwapAllowed := FALSE;
	Status.xPowerAllowed := FALSE;
	Status.xDriveResetAllowed := FALSE;
	Status.xHomeAllowed := FALSE;
	Status.xLowerAllowed := FALSE;
	Status.xRaiseAllowed := FALSE;
	Status.xSelectAllowed := FALSE;
	Status.xLockAllowed := FALSE;
	Status.xStopAllowed := FALSE;
	Status.xMoveAllowed := FALSE;
	Status.xJogAllowed := FALSE;
	Status.xTeachOperatorAllowed := FALSE;
	Status.xTeachWorkAllowed := FALSE;
	Status.xResetAllowed := FALSE;
	Status.xConfigAllowed := FALSE;
END_IF;

// Инвентарь операторской палеты редактируется всегда, независимо от режима,
// движения, подтверждения, питания и ошибок механизма. Роботная палета — только
// при выключенном магазине после освобождения текущей/выданной операции с ним,
// в том числе в Auto при работающем цикле ячейки.
// Считаем после команд и обмена, чтобы роль палеты была актуальна в этом скане.
Status.xEdit1Allowed := xSelected
	AND ((Status.uiRobotPallet <> UINT#1) OR (NOT Status.xEnabled AND xActivePalletEditAllowed));
Status.xEdit2Allowed := xSelected
	AND ((Status.uiRobotPallet <> UINT#2) OR (NOT Status.xEnabled AND xActivePalletEditAllowed));
Status.xEditAllowed := Status.xEdit1Allowed OR Status.xEdit2Allowed;
Status.xLoadAllowed := Status.xConfirmed AND NOT Status.xBusy AND NOT xOtherLoaded
	AND (((Status.uiRobotPallet = UINT#1) AND Status.xEdit2Allowed)
		OR ((Status.uiRobotPallet = UINT#2) AND Status.xEdit1Allowed));

Status.xReady := xSelected
	AND Status.xEnabled
	AND Status.xConfirmed
	AND NOT Status.xBusy
	AND NOT Status.xError
	AND xWork
	AND (uiCandidate = Status.uiRobotPallet)
	AND Input.xPowered
	AND xRobotGeometryReady
	AND xRobotMagazineReady
	AND xSafe;

IF NOT xSelected THEN
	Status.xEnabled := FALSE;
	Status.xConfirmed := FALSE;
END_IF;

(* ---- FB_TWO_PALLET_SIMULATION.st ---- *)
FUNCTION_BLOCK FB_TWO_PALLET_SIMULATION
VAR_INPUT
	xEnable : BOOL; // Только тестовая среда SIMULATION
	uiP1Signals : UINT;
	Command : ST_TWO_PALLET_OUTPUT;
END_VAR
VAR_OUTPUT
	xLiftDown : BOOL;
	xLiftUp : BOOL;
	xLockIn : BOOL;
	xLockOut : BOOL;
	xStopIn : BOOL;
	xStopOut : BOOL;
END_VAR
VAR
	xInitialized : BOOL;
	xLiftTargetUp : BOOL;
	xLockTargetOut : BOOL;
	xStopTargetOut : BOOL;
	tonLift : TON;
	tonLock : TON;
	tonStop : TON;
END_VAR

// --- BEGIN IMPLEMENTATION ---

IF NOT xEnable THEN
	xInitialized := FALSE;
	xLiftDown := FALSE;
	xLiftUp := FALSE;
	xLockIn := FALSE;
	xLockOut := FALSE;
	xStopIn := FALSE;
	xStopOut := FALSE;
	tonLift(IN := FALSE, PT := T#300MS);
	tonLock(IN := FALSE, PT := T#300MS);
	tonStop(IN := FALSE, PT := T#300MS);
ELSE
	IF NOT xInitialized THEN
		// Виртуальная начальная поза: П2 внизу, замок держит П1,
		// фиксатор держит противоположную палету.
		xLiftTargetUp := FALSE;
		xLockTargetOut := (uiP1Signals AND UINT#8) <> UINT#0;
		xStopTargetOut := (uiP1Signals AND UINT#32) <> UINT#0;
		xLiftDown := TRUE;
		xLiftUp := FALSE;
		xLockOut := xLockTargetOut;
		xLockIn := NOT xLockTargetOut;
		xStopOut := xStopTargetOut;
		xStopIn := NOT xStopTargetOut;
		xInitialized := TRUE;
	END_IF;

	// Бистабильный 5/2 сохраняет положение после снятия обеих катушек.
	IF Command.xLiftUp AND NOT Command.xLiftDown THEN
		xLiftTargetUp := TRUE;
	ELSIF Command.xLiftDown AND NOT Command.xLiftUp THEN
		xLiftTargetUp := FALSE;
	END_IF;
	IF Command.xLockOut AND NOT Command.xLockIn THEN
		xLockTargetOut := TRUE;
	ELSIF Command.xLockIn AND NOT Command.xLockOut THEN
		xLockTargetOut := FALSE;
	END_IF;
	IF Command.xStopOut AND NOT Command.xStopIn THEN
		xStopTargetOut := TRUE;
	ELSIF Command.xStopIn AND NOT Command.xStopOut THEN
		xStopTargetOut := FALSE;
	END_IF;

	tonLift(IN := xLiftTargetUp <> xLiftUp, PT := T#300MS);
	tonLock(IN := xLockTargetOut <> xLockOut, PT := T#300MS);
	tonStop(IN := xStopTargetOut <> xStopOut, PT := T#300MS);
	IF tonLift.Q THEN
		xLiftUp := xLiftTargetUp;
		xLiftDown := NOT xLiftTargetUp;
	END_IF;
	IF tonLock.Q THEN
		xLockOut := xLockTargetOut;
		xLockIn := NOT xLockTargetOut;
	END_IF;
	IF tonStop.Q THEN
		xStopOut := xStopTargetOut;
		xStopIn := NOT xStopTargetOut;
	END_IF;
END_IF;

(* ---- FB_ALARM_MANAGER.AddEvent.st ---- *)
METHOD PRIVATE AddEvent
VAR_INPUT
	eSource   : E_ALARM_SOURCE; // Источник события
	eSeverity : E_ALARM_SEVERITY; // Уровень события
	eEffect   : E_ALARM_EFFECT; // Воздействие события на ячейку
	uiCode    : UINT; // Код события внутри источника
END_VAR

// --- BEGIN IMPLEMENTATION ---

xEventsUpdated := TRUE;
udiSequence := udiSequence + 1;
IF udiSequence = UDINT#0 THEN
	udiSequence := UDINT#1;
END_IF;

Events[uiWriteIndex].udiSequence := udiSequence;
Events[uiWriteIndex].eSeverity := eSeverity;
Events[uiWriteIndex].eEffect := eEffect;
Events[uiWriteIndex].eSource := eSource;
Events[uiWriteIndex].uiCode := uiCode;
Events[uiWriteIndex].xActive := TRUE;

IF uiWriteIndex >= 100 THEN
	uiWriteIndex := 1;
ELSE
	uiWriteIndex := uiWriteIndex + 1;
END_IF;

(* ---- FB_ALARM_MANAGER.DeactivateEvent.st ---- *)
METHOD PRIVATE DeactivateEvent
VAR_INPUT
	eSource : E_ALARM_SOURCE; // Источник аварии
	uiCode  : UINT; // Номер очищенного бита
END_VAR
VAR
	uiIndex : UINT; // Индекс поиска в журнале
END_VAR

// --- BEGIN IMPLEMENTATION ---

FOR uiIndex := 1 TO 100 DO
	IF Events[uiIndex].xActive
	AND (Events[uiIndex].eSeverity = E_ALARM_SEVERITY.ALARM)
	AND (Events[uiIndex].eSource = eSource)
	AND (Events[uiIndex].uiCode = uiCode) THEN
		Events[uiIndex].xActive := FALSE;
        xEventsUpdated := TRUE;
	END_IF;
END_FOR;

(* ---- FB_ALARM_MANAGER.GetAlarmEffect.st ---- *)
METHOD PRIVATE GetAlarmEffect : E_ALARM_EFFECT
VAR_INPUT
	eSource : E_ALARM_SOURCE; // Первичный владелец ошибки
	uiCode : UINT; // Номер бита ошибки владельца
	xRobotStopRequired : BOOL; // Защёлкнутый контекст оборудования требует остановить робота
	xGlobalError : BOOL; // Активна Safety-ошибка ячейки
END_VAR

// --- BEGIN IMPLEMENTATION ---

// Safety имеет абсолютный приоритет над любой частной причиной.
IF xGlobalError THEN
	GetAlarmEffect := E_ALARM_EFFECT.GLOBAL_STOP;

ELSE
CASE eSource OF
	E_ALARM_SOURCE.CELL_SAFETY:
		GetAlarmEffect := E_ALARM_EFFECT.GLOBAL_STOP;

    E_ALARM_SOURCE.CONTROLLER_CPU_1,
    E_ALARM_SOURCE.CONTROLLER_CPU_2,
    E_ALARM_SOURCE.CONTROLLER_MODULES:
        GetAlarmEffect := E_ALARM_EFFECT.GLOBAL_STOP;

	E_ALARM_SOURCE.CELL:
		CASE uiCode OF
			1: GetAlarmEffect := E_ALARM_EFFECT.ROBOT_STOP; // ERR_ROBOT
			4: GetAlarmEffect := E_ALARM_EFFECT.GLOBAL_STOP; // ERR_GLOBAL_STOP
		ELSE GetAlarmEffect := E_ALARM_EFFECT.EQUIPMENT_STOP;
		END_CASE;

	E_ALARM_SOURCE.MACHINE_1,
	E_ALARM_SOURCE.MACHINE_2,
	E_ALARM_SOURCE.MACHINE_3:
		CASE uiCode OF
			9: GetAlarmEffect := E_ALARM_EFFECT.GLOBAL_STOP; // ERR_SAFETY_STOP
			2, 3, 13, 15, 16, 17, 23: GetAlarmEffect := E_ALARM_EFFECT.ROBOT_STOP;
		ELSE
			IF xRobotStopRequired THEN
				GetAlarmEffect := E_ALARM_EFFECT.ROBOT_STOP;
			ELSE
				GetAlarmEffect := E_ALARM_EFFECT.EQUIPMENT_STOP;
			END_IF;
		END_CASE;

	E_ALARM_SOURCE.MAGAZINE_LOGIC_1,
	E_ALARM_SOURCE.MAGAZINE_LOGIC_2:
		CASE uiCode OF
			5: GetAlarmEffect := E_ALARM_EFFECT.ROBOT_STOP; // ERR_ROBOT
			6: GetAlarmEffect := E_ALARM_EFFECT.GLOBAL_STOP; // ERR_GLOBAL_STOP
		ELSE
			IF xRobotStopRequired THEN
				GetAlarmEffect := E_ALARM_EFFECT.ROBOT_STOP;
			ELSE
				GetAlarmEffect := E_ALARM_EFFECT.EQUIPMENT_STOP;
			END_IF;
		END_CASE;

	E_ALARM_SOURCE.RESERVED_LEGACY_MAGAZINE_AXIS_1,
	E_ALARM_SOURCE.RESERVED_LEGACY_MAGAZINE_AXIS_2,
	E_ALARM_SOURCE.GEOMETRY_1,
	E_ALARM_SOURCE.GEOMETRY_2:
		IF xRobotStopRequired THEN
			GetAlarmEffect := E_ALARM_EFFECT.ROBOT_STOP;
		ELSE
			GetAlarmEffect := E_ALARM_EFFECT.EQUIPMENT_STOP;
		END_IF;

	E_ALARM_SOURCE.ROBOT,
	E_ALARM_SOURCE.AXIS_X,
	E_ALARM_SOURCE.AXIS_Y,
	E_ALARM_SOURCE.AXIS_Z,
	E_ALARM_SOURCE.AXIS_GROUP,
	E_ALARM_SOURCE.MOTION_MANAGER,
	E_ALARM_SOURCE.POINT_MANAGER,
	E_ALARM_SOURCE.GRIPPER:
		GetAlarmEffect := E_ALARM_EFFECT.ROBOT_STOP;

ELSE
	GetAlarmEffect := E_ALARM_EFFECT.EQUIPMENT_STOP;
END_CASE;
END_IF;

(* ---- FB_ALARM_MANAGER.UpdateSource.st ---- *)
METHOD PRIVATE UpdateSource
VAR_INPUT
	eSource   : E_ALARM_SOURCE; // Источник проверяемой маски ошибок
	dwCurrent : DWORD; // Текущая маска ошибок
	xRobotStopRequired : BOOL; // Контекст владельца требует зависимого останова робота
	xGlobalError : BOOL; // Глобальная ошибка активна
END_VAR
VAR_IN_OUT
	dwPrevious : DWORD; // Маска ошибок прошлого цикла
END_VAR
VAR
	dwChanged : DWORD; // Изменившиеся биты
	dwBit     : DWORD; // Маска проверяемого бита
	uiBit     : UINT; // Номер проверяемого бита
END_VAR

// --- BEGIN IMPLEMENTATION ---

dwChanged := dwCurrent XOR dwPrevious;

IF dwChanged <> DWORD#0 THEN
	FOR uiBit := 0 TO 31 DO
		dwBit := SHL(DWORD#1, uiBit);
		IF (dwChanged AND dwBit) <> DWORD#0 THEN
			IF (dwCurrent AND dwBit) <> DWORD#0 THEN
				AddEvent(
					eSource := eSource,
					eSeverity := E_ALARM_SEVERITY.ALARM,
					eEffect := GetAlarmEffect(
						eSource := eSource,
						uiCode := uiBit,
						xRobotStopRequired := xRobotStopRequired,
						xGlobalError := xGlobalError
					),
					uiCode := uiBit
				);
			ELSE
				DeactivateEvent(eSource := eSource, uiCode := uiBit);
			END_IF;
		END_IF;
	END_FOR;
	dwPrevious := dwCurrent;
END_IF;

(* ---- FB_AXIS.UpdateErrorView.st ---- *)
METHOD UpdateErrorView : ST_AXIS_ERROR
VAR_INPUT
	dwAxisError   : DWORD; // Маска ошибок SoftMotion и привода
	dwLogicalError: DWORD; // Маска логических ошибок оси
END_VAR
VAR
	stError : ST_AXIS_ERROR; // Представление ошибок отдельными флагами
END_VAR

// --- BEGIN IMPLEMENTATION ---

stError.MC_POWER_ERROR := (dwAxisError AND AXE_MC_POWER_ERROR) <> DWORD#0;
stError.MC_RESET_ERROR := (dwAxisError AND AXE_MC_RESET_ERROR) <> DWORD#0;
stError.MC_STOP_ERROR := (dwAxisError AND AXE_MC_STOP_ERROR) <> DWORD#0;
stError.MC_JOG_ERROR := (dwAxisError AND AXE_MC_JOG_ERROR) <> DWORD#0;
stError.MC_HOME_ERROR := (dwAxisError AND AXE_MC_HOME_ERROR) <> DWORD#0;
stError.MC_MOVE_ABS_ERROR := (dwAxisError AND AXE_MC_MOVE_ABS_ERROR) <> DWORD#0;
stError.MC_MOVE_REL_ERROR := (dwAxisError AND AXE_MC_MOVE_REL_ERROR) <> DWORD#0;
stError.READ_POSITION_ERROR := (dwAxisError AND AXE_READ_POS_ERROR) <> DWORD#0;
stError.READ_STATUS_ERROR := (dwAxisError AND AXE_READ_STATUS_ERROR) <> DWORD#0;
stError.AXIS_ERRORSTOP := (dwAxisError AND AXE_ERRORSTOP) <> DWORD#0;
stError.FB_ERROR_OCCURRED := (dwAxisError AND AXE_FB_ERROR_OCCURRED) <> DWORD#0;
stError.COMMAND_ABORTED := (dwAxisError AND AXE_COMMAND_ABORTED) <> DWORD#0;
stError.UNKNOWN_AXIS_ERROR := (dwAxisError AND AXE_UNKNOWN_ACTUAL_ERROR) <> DWORD#0;
stError.DRIVE_AXIS_ERROR := (dwAxisError AND AXE_DRIVE_AXIS_ERROR) <> DWORD#0;
stError.POWER_FEEDBACK_LOST := (dwAxisError AND AXE_POWER_FEEDBACK_LOST) <> DWORD#0;

stError.POWER_PERMIT_LOST := (dwLogicalError AND LOG_POWER_PERMIT_LOST) <> DWORD#0;
stError.GLOBAL_DURING_POWER := (dwLogicalError AND LOG_GLOBAL_DURING_POWER) <> DWORD#0;
stError.GLOBAL_DURING_READY := (dwLogicalError AND LOG_GLOBAL_DURING_READY) <> DWORD#0;
stError.GLOBAL_DURING_MOTION := (dwLogicalError AND LOG_GLOBAL_DURING_MOTION) <> DWORD#0;
stError.JOG_CONFLICT := (dwLogicalError AND LOG_JOG_CONFLICT) <> DWORD#0;
stError.MOVE_ABS_NOT_HOMED := (dwLogicalError AND LOG_MOVE_ABS_NOT_HOMED) <> DWORD#0;
stError.MOVE_REL_NOT_HOMED := (dwLogicalError AND LOG_MOVE_REL_NOT_HOMED) <> DWORD#0;
stError.STEP_TIMEOUT := (dwLogicalError AND LOG_STEP_TIMEOUT) <> DWORD#0;
stError.UNKNOWN_STEP := (dwLogicalError AND LOG_UNKNOWN_STEP) <> DWORD#0;

UpdateErrorView := stError;

(* ---- FB_AXIS_GROUP.UpdateErrorView.st ---- *)
METHOD UpdateErrorView : ST_AXIS_GROUP_ERROR
VAR_INPUT
	dwMotionError : DWORD; // Маска ошибок блоков SoftMotion
	dwLogicalError: DWORD; // Маска логических ошибок группы
END_VAR
VAR
	stError : ST_AXIS_GROUP_ERROR; // Представление ошибок отдельными флагами
END_VAR

// --- BEGIN IMPLEMENTATION ---

stError.ENABLE_ERROR := (dwMotionError AND MOTION_ERR_ENABLE) <> DWORD#0;
// Зарезервировано для совместимости символов: питанием осей владеют FB_AXIS.
stError.POWER_ERROR := FALSE;
stError.DISABLE_ERROR := (dwMotionError AND MOTION_ERR_DISABLE) <> DWORD#0;
stError.RESET_ERROR := (dwMotionError AND MOTION_ERR_RESET) <> DWORD#0;
stError.MOVE_DIRECT_ERROR := (dwMotionError AND MOTION_ERR_MOVE_DIRECT) <> DWORD#0;
stError.MOVE_LINEAR_ERROR := (dwMotionError AND MOTION_ERR_MOVE_LINEAR) <> DWORD#0;
stError.HALT_ERROR := (dwMotionError AND MOTION_ERR_HALT) <> DWORD#0;
stError.STOP_ERROR := (dwMotionError AND MOTION_ERR_STOP) <> DWORD#0;
stError.READ_POSITION_ERROR := (dwMotionError AND MOTION_ERR_READ_POSITION) <> DWORD#0;
stError.READ_STATUS_ERROR := (dwMotionError AND MOTION_ERR_READ_STATUS) <> DWORD#0;
stError.READ_GROUP_ERROR := (dwMotionError AND MOTION_ERR_READ_GROUP_ERROR) <> DWORD#0;
stError.GROUP_ERROR_STOP := (dwMotionError AND MOTION_ERR_GROUP_ERROR_STOP) <> DWORD#0;
stError.SIMULATED_ERROR := (dwMotionError AND MOTION_ERR_SIMULATED) <> DWORD#0;
stError.OVERRIDE_ERROR := (dwMotionError AND MOTION_ERR_OVERRIDE) <> DWORD#0;

stError.STEP_TIMEOUT := (dwLogicalError AND LOG_STEP_TIMEOUT) <> DWORD#0;
stError.INVALID_STATE := (dwLogicalError AND LOG_INVALID_STATE) <> DWORD#0;
stError.POWER_PERMIT_READY := (dwLogicalError AND LOG_POWER_PERMIT_READY) <> DWORD#0;
stError.POWER_PERMIT_LOST := (dwLogicalError AND LOG_POWER_PERMIT_LOST_DIRECT) <> DWORD#0;

UpdateErrorView := stError;

(* ---- FB_CELL_SAFETY.RaiseWarning.st ---- *)
METHOD PRIVATE RaiseWarning
VAR_INPUT
	uiCode : UINT;
END_VAR

// --- BEGIN IMPLEMENTATION ---

Diag.stWarning.uiCode := uiCode;
Diag.stWarning.udiSequence := Diag.stWarning.udiSequence + UDINT#1;
IF Diag.stWarning.udiSequence = UDINT#0 THEN
	Diag.stWarning.udiSequence := UDINT#1;
END_IF;

(* ---- FB_GRIPPER_SIMULATION.UpdateErrorView.st ---- *)
METHOD UpdateErrorView : ST_GRIPPER_ERROR
VAR_INPUT
	dwError : DWORD; // Битовая маска для расшифровки
END_VAR
VAR
	stError : ST_GRIPPER_ERROR; // Представление ошибок отдельными флагами
END_VAR

// --- BEGIN IMPLEMENTATION ---

stError.GRIPPER_1_ERROR := (dwError AND ERR_GRIPPER_1) <> DWORD#0;
stError.GRIPPER_2_ERROR := (dwError AND ERR_GRIPPER_2) <> DWORD#0;
stError.ROTATION_ERROR := (dwError AND ERR_GRIP_ROTATE) <> DWORD#0;
stError.ACTION_ERROR := (dwError AND ERR_GRIP_ACTION) <> DWORD#0;
stError.GLOBAL_ERROR := (dwError AND ERR_GRIP_GLOBAL) <> DWORD#0;

UpdateErrorView := stError;

(* ---- FB_MACHINE.UpdateErrorView.st ---- *)
METHOD UpdateErrorView : ST_MACHINE_ERROR
VAR_INPUT
	dwError : DWORD; // Битовая маска для расшифровки
END_VAR
VAR
	stError : ST_MACHINE_ERROR; // Представление ошибок отдельными флагами
END_VAR

// --- BEGIN IMPLEMENTATION ---

stError.WRONG_OPERATION := (dwError AND ERR_WRONG_OPERATION) <> DWORD#0;
stError.WRONG_COMMAND := (dwError AND ERR_WRONG_COMMAND) <> DWORD#0;
stError.ROBOT_MOTION := (dwError AND ERR_ROBOT_MOTION) <> DWORD#0;
stError.ROBOT_ACTION := (dwError AND ERR_ROBOT_ACTION) <> DWORD#0;
stError.DOOR_OPEN := (dwError AND ERR_DOOR_OPEN) <> DWORD#0;
stError.DOOR_CLOSE := (dwError AND ERR_DOOR_CLOSE) <> DWORD#0;
stError.CHUCK_OPEN := (dwError AND ERR_CHUCK_OPEN) <> DWORD#0;
stError.CHUCK_CLOSE := (dwError AND ERR_CHUCK_CLOSE) <> DWORD#0;
stError.CYCLE_START := (dwError AND ERR_CYCLE_START) <> DWORD#0;
stError.SAFETY_STOP := (dwError AND ERR_SAFETY_STOP) <> DWORD#0;
stError.UNKNOWN_DETAIL := (dwError AND ERR_UNKNOWN_DETAIL) <> DWORD#0;
stError.MACHINE_ALARM := (dwError AND ERR_MACHINE_ALARM) <> DWORD#0;
stError.INDEX_ERROR := (dwError AND ERR_INDEX) <> DWORD#0;
stError.DOOR_ROBOT := (dwError AND ERR_DOOR_ROBOT) <> DWORD#0;
stError.MACHINE_IDLE := (dwError AND ERR_MACHINE_IDLE) <> DWORD#0;
stError.TIMEOUT_ROBOT_MOVE := (dwError AND ERR_TIMEOUT_ROBOT_MOVE) <> DWORD#0;
stError.TIMEOUT_ROBOT_ACTION := (dwError AND ERR_TIMEOUT_ROBOT_ACTION) <> DWORD#0;
stError.TIMEOUT_ROBOT_RELEASE := (dwError AND ERR_TIMEOUT_ROBOT_RELEASE) <> DWORD#0;
stError.TIMEOUT_DOOR_OPEN := (dwError AND ERR_TIMEOUT_DOOR_OPEN) <> DWORD#0;
stError.TIMEOUT_DOOR_CLOSE := (dwError AND ERR_TIMEOUT_DOOR_CLOSE) <> DWORD#0;
stError.TIMEOUT_HATCH_UNLOCK := (dwError AND ERR_TIMEOUT_HATCH_UNLOCK) <> DWORD#0;
stError.TIMEOUT_CHUCK_OPEN := (dwError AND ERR_TIMEOUT_CHUCK_OPEN) <> DWORD#0;
stError.TIMEOUT_CHUCK_CLOSE := (dwError AND ERR_TIMEOUT_CHUCK_CLOSE) <> DWORD#0;
stError.TIMEOUT_CYCLE_START := (dwError AND ERR_TIMEOUT_CYCLE_START) <> DWORD#0;
stError.SAFETY_DOOR_OPEN := (dwError AND ERR_SAFETY_DOOR_OPEN) <> DWORD#0;
stError.HATCH_UNLOCK_PROCESSING := (dwError AND ERR_HATCH_UNLOCK_PROCESSING) <> DWORD#0;

UpdateErrorView := stError;

(* ---- FB_MACHINE_SIMULATION.UpdateErrorView.st ---- *)
METHOD UpdateErrorView : ST_MACHINE_SIM_ERROR
VAR_INPUT
	dwError : DWORD; // Битовая маска для расшифровки
END_VAR
VAR
	stError : ST_MACHINE_SIM_ERROR; // Представление ошибок отдельными флагами
END_VAR

// --- BEGIN IMPLEMENTATION ---

stError.MACHINE_ALARM := (dwError AND ERR_MACHINE_ALARM) <> DWORD#0;
stError.DOOR_FAULT := (dwError AND ERR_DOOR_FAULT) <> DWORD#0;
stError.CHUCK_FAULT := (dwError AND ERR_CHUCK_FAULT) <> DWORD#0;

UpdateErrorView := stError;

(* ---- FB_MAGAZINE.FindBlank.st ---- *)
METHOD FindBlank : SINT
VAR_INPUT
	iSlotCount : SINT; // Число слотов, участвующих в поиске
END_VAR
VAR_IN_OUT
	stDetail : ARRAY [1..GVL_CELL_SETTINGS.NumberDetail] OF ST_DETAIL; // Содержимое слотов магазина
END_VAR
VAR
	i : SINT; // Индекс проверяемого слота
END_VAR

// --- BEGIN IMPLEMENTATION ---

FindBlank := 0;

FOR i:= 1 TO iSlotCount DO
	IF stDetail[i].xInPosition = TRUE AND stDetail[i].eDetailType =  E_DETAIL_TYPE.BLANK THEN
		FindBlank := i;
		EXIT;
	END_IF
END_FOR

(* ---- FB_MAGAZINE.FindFreeSlot.st ---- *)
METHOD FindFreeSlot : SINT
VAR_INPUT
	iSlotCount : SINT; // Число слотов, участвующих в поиске
END_VAR
VAR_IN_OUT
	stDetail : ARRAY [1..GVL_CELL_SETTINGS.NumberDetail] OF ST_DETAIL; // Содержимое слотов магазина
END_VAR
VAR
	i : SINT; // Индекс проверяемого слота
END_VAR

// --- BEGIN IMPLEMENTATION ---

FindFreeSlot := 0;

FOR i:= 1 TO iSlotCount DO
	IF stDetail[i].xInPosition = FALSE THEN
		FindFreeSlot := i;
		EXIT;
	END_IF
END_FOR

(* ---- FB_MAGAZINE.UpdateErrorView.st ---- *)
METHOD UpdateErrorView : ST_MAGAZINE_ERROR
VAR_INPUT
	dwError : DWORD; // Битовая маска для расшифровки
END_VAR
VAR
	stError : ST_MAGAZINE_ERROR; // Представление ошибок отдельными флагами
END_VAR

// --- BEGIN IMPLEMENTATION ---

stError.WRONG_OPERATION := (dwError AND ERR_WRONG_OPERATION) <> DWORD#0;
stError.NO_BLANK := (dwError AND ERR_NO_BLANK) <> DWORD#0;
stError.NO_FREE_SLOT := (dwError AND ERR_NO_FREE_SLOT) <> DWORD#0;
stError.INVALID_SLOT := (dwError AND ERR_INVALID_SLOT) <> DWORD#0;
stError.SLOT_CONTENT := (dwError AND ERR_SLOT_CONTENT) <> DWORD#0;
stError.ROBOT_ERROR := (dwError AND ERR_ROBOT) <> DWORD#0;
stError.GLOBAL_STOP := (dwError AND ERR_GLOBAL_STOP) <> DWORD#0;
stError.GEOMETRY_ERROR := (dwError AND ERR_GEOMETRY) <> DWORD#0;

UpdateErrorView := stError;

(* ---- FB_MAGAZINE.UpdateTypeStatus.st ---- *)
METHOD PRIVATE UpdateTypeStatus
VAR_IN_OUT
    stMagazineInventory : ST_MAGAZINE_INVENTORY;
END_VAR
VAR
    uiType : UINT;
    uiSlot : UINT;
    iSlot : SINT;
    uiFreeCount : UINT;
    xValidTypeCount : BOOL;
END_VAR

// --- BEGIN IMPLEMENTATION ---

// Один проход даёт выбор слотов и сводку. Пустое место универсально для типов.
iInventoryFirstBlank := SINT#0;
iInventoryFirstFree := SINT#0;
uiFreeCount := UINT#0;
xValidTypeCount := (uiTypeCount >= UINT#1) AND (uiTypeCount <= UINT#3);
FOR uiType := UINT#1 TO UINT#3 DO
    Status.stTypeStatus.aiBlankSlot[uiType] := SINT#0;
    Status.stTypeStatus.aiFreeSlot[uiType] := SINT#0;
    Status.stTypeStatus.auiBlankCount[uiType] := UINT#0;
    Status.stTypeStatus.auiDetailCount[uiType] := UINT#0;
    Status.stTypeStatus.auiFreeCount[uiType] := UINT#0;
END_FOR;
IF iActiveSlotCount > SINT#0 THEN
    FOR uiSlot := UINT#1 TO SINT_TO_UINT(iActiveSlotCount) DO
        iSlot := UINT_TO_SINT(uiSlot);
        IF NOT stMagazineInventory.aSlots[iSlot].xInPosition THEN
            uiFreeCount := uiFreeCount + UINT#1;
            IF iInventoryFirstFree = SINT#0 THEN iInventoryFirstFree := iSlot; END_IF;
        ELSE
            IF (iInventoryFirstBlank = SINT#0)
            AND (stMagazineInventory.aSlots[iSlot].eDetailType = E_DETAIL_TYPE.BLANK) THEN
                iInventoryFirstBlank := iSlot;
            END_IF;
            uiType := stMagazineInventory.aSlots[iSlot].uiProductType;
            IF xValidTypeCount AND (uiType >= UINT#1) AND (uiType <= uiTypeCount) THEN
                IF stMagazineInventory.aSlots[iSlot].eDetailType = E_DETAIL_TYPE.BLANK THEN
                    Status.stTypeStatus.auiBlankCount[uiType] := Status.stTypeStatus.auiBlankCount[uiType] + UINT#1;
                    IF Status.stTypeStatus.aiBlankSlot[uiType] = SINT#0 THEN Status.stTypeStatus.aiBlankSlot[uiType] := iSlot; END_IF;
                ELSIF stMagazineInventory.aSlots[iSlot].eDetailType = E_DETAIL_TYPE.DETAIL THEN
                    Status.stTypeStatus.auiDetailCount[uiType] := Status.stTypeStatus.auiDetailCount[uiType] + UINT#1;
                END_IF;
            END_IF;
        END_IF;
    END_FOR;
END_IF;
IF xValidTypeCount THEN
    FOR uiType := UINT#1 TO uiTypeCount DO
        Status.stTypeStatus.auiFreeCount[uiType] := uiFreeCount;
        Status.stTypeStatus.aiFreeSlot[uiType] := iInventoryFirstFree;
    END_FOR;
END_IF;
iInventorySummarySlotCount := iActiveSlotCount;
uiInventorySummaryTypeCount := uiTypeCount;
xInventorySummaryInitialized := TRUE;
xInventorySummaryDirty := FALSE;

(* ---- FB_MOTION_MANAGER.UpdateErrorView.st ---- *)
METHOD UpdateErrorView : ST_MOTION_MANAGER_ERROR
VAR_INPUT
	dwError : DWORD; // Битовая маска для расшифровки
END_VAR
VAR
	stError : ST_MOTION_MANAGER_ERROR; // Представление ошибок отдельными флагами
END_VAR

// --- BEGIN IMPLEMENTATION ---

stError.POINT_INVALID := (dwError AND ERR_POINT_INVALID) <> DWORD#0;
stError.GROUP_ERROR := (dwError AND ERR_GROUP) <> DWORD#0;
stError.GLOBAL_STOP := (dwError AND ERR_GLOBAL_STOP) <> DWORD#0;
stError.START_TIMEOUT := (dwError AND ERR_START_TIMEOUT) <> DWORD#0;

UpdateErrorView := stError;

(* ---- FB_POINT_MANAGER.UpdateErrorView.st ---- *)
METHOD UpdateErrorView : ST_POINT_MANAGER_ERROR
VAR_INPUT
	dwError : DWORD; // Битовая маска для расшифровки
END_VAR
VAR
	stError : ST_POINT_MANAGER_ERROR; // Представление ошибок отдельными флагами
END_VAR

// --- BEGIN IMPLEMENTATION ---

stError.X_OUT_OF_LIMIT := (dwError AND X_OUT_OF_LIMIT) <> DWORD#0;
stError.Y_OUT_OF_LIMIT := (dwError AND Y_OUT_OF_LIMIT) <> DWORD#0;
stError.Z_OUT_OF_LIMIT := (dwError AND Z_OUT_OF_LIMIT) <> DWORD#0;
stError.INVALID_VEL := (dwError AND INVALID_VEL) <> DWORD#0;
stError.X_LIMIT_CONFIG_INVALID := (dwError AND X_LIMIT_CONFIG_INVALID) <> DWORD#0;
stError.Y_LIMIT_CONFIG_INVALID := (dwError AND Y_LIMIT_CONFIG_INVALID) <> DWORD#0;
stError.Z_LIMIT_CONFIG_INVALID := (dwError AND Z_LIMIT_CONFIG_INVALID) <> DWORD#0;
stError.POINT_NOT_CONFIGURED := (dwError AND POINT_NOT_CONFIGURED) <> DWORD#0;

UpdateErrorView := stError;

(* ---- FB_ROBOT.UpdateErrorView.st ---- *)
METHOD UpdateErrorView : ST_ROBOT_ERROR
VAR_INPUT
	dwError : DWORD; // Битовая маска для расшифровки
END_VAR
VAR
	stError : ST_ROBOT_ERROR; // Представление ошибок отдельными флагами
END_VAR

// --- BEGIN IMPLEMENTATION ---

stError.WRONG_ACTION := (dwError AND ERR_ROBOT_WRONG_ACTION) <> DWORD#0;
stError.MOTION_ERROR := (dwError AND ERR_ROBOT_MOTION) <> DWORD#0;
stError.GRIPPER_ERROR := (dwError AND ERR_ROBOT_GRIPPER) <> DWORD#0;
stError.MODBUS_COMMUNICATION_ERROR := (dwError AND ERR_ROBOT_MODBUS_COMM) <> DWORD#0;
stError.EXTERNAL_ROBOT_ALARM := (dwError AND ERR_EXTERNAL_ROBOT) <> DWORD#0;
stError.MODBUS_ERROR := stError.MODBUS_COMMUNICATION_ERROR OR stError.EXTERNAL_ROBOT_ALARM;
stError.STOP_ERROR := (dwError AND ERR_ROBOT_STOP) <> DWORD#0;

UpdateErrorView := stError;

(* ---- FB_TWO_PALLET.IsSignalConfigurationValid.st ---- *)
METHOD IsSignalConfigurationValid : BOOL
VAR_INPUT
	uiP1Signals : UINT;
	uiP2Signals : UINT;
END_VAR

// --- BEGIN IMPLEMENTATION ---

// Рабочее положение каждого цилиндра подтверждает ровно один геркон.
// Зацепление должно различать палеты и при опущенной П2 во время обмена.
IsSignalConfigurationValid := (uiP1Signals <= UINT#63)
	AND (uiP2Signals <= UINT#63)
	AND (((uiP1Signals AND UINT#3) = UINT#1) OR ((uiP1Signals AND UINT#3) = UINT#2))
	AND (((uiP2Signals AND UINT#3) = UINT#1) OR ((uiP2Signals AND UINT#3) = UINT#2))
	AND (((uiP1Signals AND UINT#12) = UINT#4) OR ((uiP1Signals AND UINT#12) = UINT#8))
	AND (((uiP2Signals AND UINT#12) = UINT#4) OR ((uiP2Signals AND UINT#12) = UINT#8))
	AND (((uiP1Signals AND UINT#48) = UINT#16) OR ((uiP1Signals AND UINT#48) = UINT#32))
	AND (((uiP2Signals AND UINT#48) = UINT#16) OR ((uiP2Signals AND UINT#48) = UINT#32))
	AND ((uiP1Signals AND UINT#60) <> (uiP2Signals AND UINT#60));

(* ---- FB_TWO_PALLET.UpdateErrorView.st ---- *)
METHOD UpdateErrorView : ST_TWO_PALLET_ERROR
VAR_INPUT
	dwError : DWORD;
END_VAR
VAR
	stError : ST_TWO_PALLET_ERROR;
END_VAR

// --- BEGIN IMPLEMENTATION ---

stError.DRIVE_ERROR := (dwError AND ERR_DRIVE) <> DWORD#0;
stError.SENSOR_CONTRADICTION := (dwError AND ERR_SENSOR_CONTRADICTION) <> DWORD#0;
stError.CYLINDER_TIMEOUT := (dwError AND ERR_CYLINDER_TIMEOUT) <> DWORD#0;
stError.MOTION_TIMEOUT := (dwError AND ERR_MOTION_TIMEOUT) <> DWORD#0;
stError.LOGIC_ERROR := (dwError AND ERR_LOGIC) <> DWORD#0;
stError.SEQUENCE_INTERRUPTED := (dwError AND ERR_SEQUENCE_INTERRUPTED) <> DWORD#0;

UpdateErrorView := stError;
